(*
SPDX-License-Identifier: MIT
License: https://opensource.org/license/mit
*)

(*!
<summary>Runs a valid empty root array without synthetic test results.</summary>
<description>
Owns persistent root instances and fixed child storage. Use from one task without reentry.
Children borrows the same array for the instance lifetime. Root parents remain zero.
</description>
*)

{attribute 'no_assign'}
{attribute 'no_explicit_call' := 'do not call this function block directly'}
FUNCTION_BLOCK EmptyTestRunner EXTENDS TOF_Testing.TestRunner<0>
VAR_STAT
	//! <summary>Class name shared by instances of this concrete runner.</summary>
	{attribute 'hide'}
	_ClassName : STRING := __POUNAME();
END_VAR
VAR
	{attribute 'hide'}
	{attribute 'init_namespace'}
	_NamespaceName : STRING;
END_VAR
VAR
	_Children : ARRAY [0.._ChildCount - 1] OF TOF_Testing.ITestElement;
END_VAR

(*!
<summary>Borrows the concrete class name; callers must not modify the returned storage.</summary>
*)
{attribute 'monitoring' := 'call'}
PROPERTY ClassName : REFERENCE TO STRING
GET
ClassName REF= _ClassName;
END_GET
END_PROPERTY

(*!
<summary>Borrows the concrete namespace name for the instance lifetime; callers must not modify it.</summary>
*)
{attribute 'monitoring' := 'call'}
PROPERTY NamespaceName : REFERENCE TO STRING
GET
NamespaceName REF= _NamespaceName;
END_GET
END_PROPERTY

(*!
<summary>Reports the complete concrete instance size.</summary>
*)
{attribute 'monitoring' := 'call'}
PROPERTY SelfSize : ULINT
GET
SelfSize := XSIZEOF(THIS^);
END_GET
END_PROPERTY

(*!
<summary>Borrows the unchanged persistent root array; application code must not modify it.</summary>
*)
{attribute 'monitoring' := 'call'}
PROPERTY Children : REFERENCE TO ARRAY [0.._ChildCount - 1] OF TOF_Testing.ITestElement
GET
Children REF= _Children;
END_GET
END_PROPERTY

END_FUNCTION_BLOCK

(* stored: Version 1.1.0.1
   POU EmptyTestRunner: Id {c0097876-f043-4e94-b0ea-9af4f803ccae}, SpecialFunc None
   Property ClassName: Id {13d1f45e-0875-44ea-9267-9ea0102be582}
   Get Get: Id {75b02eed-cb92-4bf2-bea7-a35baf4316e4}
   Property NamespaceName: Id {4c11365b-e099-41f4-8f82-98fb7deecd13}
   Get Get: Id {0607d826-0e9e-44f1-9d5e-0e421310c660}
   Property SelfSize: Id {8486738b-ac87-4908-9947-8a79aa1237d4}
   Get Get: Id {e8d276a9-24a3-44d9-9246-9a6d0f0f237d}
   Property Children: Id {286bbd78-2e5e-4d8c-ac24-f87048191b9b}
   Get Get: Id {f42b0288-bc03-479b-9bef-2239600a8be3} *)
